// TIA Portal V21 export
// export: Created 2026-10-14T03:09:04.8839945Z, ExportSetting WithDefaults, DisplayName Totally Integrated Automation Portal, DisplayVersion V21, DisplayName STEP 7 Professional, DisplayVersion V21, DisplayName STEP 7 Safety, DisplayVersion V21, DisplayName Tech WebApplication, DisplayVersion V21, DisplayName WinCC Basic/Comfort/Advanced, DisplayVersion V21, DisplayName WinCC Unified, DisplayVersion V21
Screen "10_Startscreen"  800x480, Number=18, Template=01_One_Nav_Level
  on GenerateScreen: GetStartScreenName(); SetTag(Tag := MainNavigationState, Value := 1)
  ScreenLayer 
    Button "Button_12" at 45,392 size 90x32  Mode=Text, TextOff="Place bottle", TextOn="Place bottles"
      VisibilityAnimation "VisibilityAnimation"  RangeEnd=1, RangeStart=1
        tag hmiError
      on Press: ResetBit(Tag := hmiError)
    Rectangle "Rectangle_8" at 682,361 size 88x104  StyleItem=Rectangle
      VisibilityAnimation "VisibilityAnimation"  RangeEnd=1, RangeStart=1
        tag HMI_bottleInfoActive
    GraphicView "Graphic view_4" at 213,87 size 249x237  Picture=Graphic_13
    Button "Button_4" at 45,159 size 90x48  Mode=Text, TextOff="Start", TextOn="Text"
      RangeAppearanceAnimation "RangeAppearanceAnimation"
        tag stateRunning
        0..0: back #404d53, fore #ffffff
      ObjectEnablingAnimation "ObjectEnablingAnimation"
        tag stateRunning
      on Press: SetBit(Tag := hmiStart)
      on Release: ResetBit(Tag := hmiStart)
    Button "Button_5" at 45,215 size 90x48  Mode=Text, TextOff="Stop", TextOn="Text"
      RangeAppearanceAnimation "RangeAppearanceAnimation"
        tag stateRunning
        1..1: back #404d53, fore #ffffff
      ObjectEnablingAnimation "ObjectEnablingAnimation"  RangeEnd=1, RangeStart=1
        tag stateRunning
      on Press: SetBit(Tag := hmiStop)
      on Release: ResetBit(Tag := hmiStop)
    Button "Button_6" at 45,271 size 90x48  Mode=Text, TextOff="Reset", TextOn="Text"
      RangeAppearanceAnimation "RangeAppearanceAnimation"
        tag stateStop
        1..1: back #404d53, fore #ffffff
      ObjectEnablingAnimation "ObjectEnablingAnimation"  RangeEnd=1, RangeStart=1
        tag stateStop
      on Press: SetBit(Tag := hmiReset); ResetBit(Tag := HMI_bottleInfo1); ResetBit(Tag := HMI_bottleInfo2); ResetBit(Tag := HMI_bottleInfo3); ResetBit(Tag := HMI_bottleInfo4); ResetBit(Tag := HMI_bottleInfoActive)
      on Release: ResetBit(Tag := hmiReset)
    IOField "ioKPI" at 700,269 size 68x28  DataFormat=Decimal, FormatPattern=99.9, Mode=Output
      ProcessValue := tankTemperature
    IOField "ioKPI_1" at 687,239 size 76x28  DataFormat=Decimal, FormatPattern=9999, Mode=Output
      ProcessValue := tankLevel
    TextField "Text field_3" at 496,160 size 150x25  Text="Bottles produced"
    Button "Button_1" at 45,354 size 90x32  Mode=Text, TextOff="Next bottle", TextOn="Text"
      ObjectEnablingAnimation "ObjectEnablingAnimation"  RangeEnd=1, RangeStart=1
        tag stateFillingBottle
      RangeAppearanceAnimation "RangeAppearanceAnimation"
        tag stateFillingBottle
        1..1: back #404d53, fore #ffffff
      on Press: SetBit(Tag := hmiNextBottle)
      on Release: ResetBit(Tag := hmiNextBottle)
    TextField "Text field_1" at 610,106 size 150x25  Text="Filling tank"
      VisibilityAnimation "VisibilityAnimation"  Visible=false
        tag stateFillingTank
    TextField "Text field_5" at 496,106 size 49x25  Text="State"
    TextField "Text field_6" at 610,106 size 150x25  Text="Heating tank"
      VisibilityAnimation "VisibilityAnimation"  Visible=false
        tag stateHeatingTank
    TextField "Text field_7" at 610,106 size 150x25  Text="Filling bottle"
      VisibilityAnimation "VisibilityAnimation"  Visible=false
        tag stateFillingBottle
    TextField "Text field_8" at 610,106 size 150x25  Text="Shifting bottle"
      VisibilityAnimation "VisibilityAnimation"  Visible=false
        tag stateShiftingBottle
    TextField "Text field_9" at 610,106 size 150x25  Text="Stop"
      VisibilityAnimation "VisibilityAnimation"  Visible=false
        tag stateStop
    TextField "Text field_10" at 610,106 size 150x25  Text="Reset"
      VisibilityAnimation "VisibilityAnimation"  Visible=false
        tag stateReset
    IOField "ioKPI_2" at 638,160 size 124x28  DataFormat=Decimal, FormatPattern=9999999999, Mode=Output
      ProcessValue := bottlesProduced
    TextField "Text field_11" at 496,191 size 119x25  Text="Bottles faulty"
    IOField "ioKPI_3" at 638,191 size 124x28  DataFormat=Decimal, FormatPattern=9999999999, Mode=Output
      ProcessValue := bootleNumberFaulty
    IOField "ioKPI_4" at 695,329 size 68x28  DataFormat=Decimal, FormatPattern=9.99, Mode=Output
      ProcessValue := bottleLevel
    GraphicView "Graphic view_13" at 326,321 size 17x21  Picture=Graphic_18
    Bar "Bar_1" at 223,115 size 229x206  CountSubDivisions=5, IntegerDigits=3, LargeTickLabelingStep=2, MaximumValue=1600
      RangeAppearanceAnimation "RangeAppearanceAnimation"
        tag tankTemperature
        30..39: back #adaeb5, fore #3f3cff
        40..49: back #adaeb5, fore #4f4dff
        50..59: back #adaeb5, fore #4f4dff
        60..69: back #adaeb5, fore #605eff
        70..72: back #adaeb5, fore #716eff
        73..74: back #adaeb5, fore #8280ff
        75..75: back #adaeb5, fore #9291ff
        76..76: back #adaeb5, fore #9291ff
        77..77: back #adaeb5, fore #a3a2ff
        78..78: back #adaeb5, fore #a3a2ff
        79..79: back #adaeb5, fore #b4b2ff
        80..100: back #adaeb5, fore #b4b2ff
      ProcessValue := tankLevel
    GraphicView "Graphic view_7" at 617,192 size 23x23  Picture=Graphic_58
      VisibilityAnimation "VisibilityAnimation"  RangeEnd=1, RangeStart=1
        tag bottleFaulty
    Rectangle "Rectangle_1" at 238,418 size 32x8  StyleItem=Rectangle
    Rectangle "Rectangle_2" at 199,418 size 32x8  StyleItem=Rectangle
    Line "Line_1" at 200,422 size 266x0  StyleItem=Line
      VisibilityAnimation "VisibilityAnimation"  RangeEnd=2, Visible=false
        tag bottlesProduced
    Rectangle "Rectangle_3" at 279,418 size 32x8  StyleItem=Rectangle
    Rectangle "Rectangle_4" at 317,418 size 32x8  StyleItem=Rectangle
    Rectangle "Rectangle_5" at 356,418 size 32x8  StyleItem=Rectangle
      VisibilityAnimation "VisibilityAnimation"  Visible=false
        tag bottlesProduced
    Rectangle "Rectangle_6" at 396,418 size 32x8  StyleItem=Rectangle
      VisibilityAnimation "VisibilityAnimation"  RangeEnd=1, Visible=false
        tag bottlesProduced
    Rectangle "Rectangle_7" at 436,418 size 32x8  StyleItem=Rectangle
      VisibilityAnimation "VisibilityAnimation"  RangeEnd=2, Visible=false
        tag bottlesProduced
    Line "Line_2" at 200,422 size 225x0  StyleItem=Line
      VisibilityAnimation "VisibilityAnimation"  RangeEnd=1, Visible=false
        tag bottlesProduced
    Line "Line_3" at 200,422 size 185x0  StyleItem=Line
      VisibilityAnimation "VisibilityAnimation"  Visible=false
        tag bottlesProduced
    Line "Line_4" at 201,422 size 147x0  StyleItem=Line
    Button "Button_2" at 322,431 size 26x22  Mode=Graphic, PictureOff=Graphic_50, StyleItem=Button, TextOff="Text", TextOn="Text"
      on Click: SetBit(Tag := HMI_bottleInfo1); ResetBit(Tag := HMI_bottleInfo2); ResetBit(Tag := HMI_bottleInfo3); ResetBit(Tag := HMI_bottleInfo4); HandleBottleInfo()
    Button "Button_7" at 361,431 size 26x22  Mode=Graphic, PictureOff=Graphic_50, StyleItem=Button, TextOff="Text", TextOn="Text"
      VisibilityAnimation "VisibilityAnimation"  Visible=false
        tag bottlesProduced
      on Click: SetBit(Tag := HMI_bottleInfo2); ResetBit(Tag := HMI_bottleInfo1); ResetBit(Tag := HMI_bottleInfo3); ResetBit(Tag := HMI_bottleInfo4); HandleBottleInfo()
    Button "Button_3" at 400,431 size 26x22  Mode=Graphic, PictureOff=Graphic_50, StyleItem=Button, TextOff="Text", TextOn="Text"
      VisibilityAnimation "VisibilityAnimation"  RangeEnd=1, Visible=false
        tag bottlesProduced
      on Click: SetBit(Tag := HMI_bottleInfo3); ResetBit(Tag := HMI_bottleInfo1); ResetBit(Tag := HMI_bottleInfo2); ResetBit(Tag := HMI_bottleInfo4); HandleBottleInfo()
    Button "Button_8" at 440,430 size 26x22  Mode=Graphic, PictureOff=Graphic_50, StyleItem=Button, TextOff="Text", TextOn="Text"
      VisibilityAnimation "VisibilityAnimation"  RangeEnd=2, Visible=false
        tag bottlesProduced
      on Click: SetBit(Tag := HMI_bottleInfo4); ResetBit(Tag := HMI_bottleInfo1); ResetBit(Tag := HMI_bottleInfo2); ResetBit(Tag := HMI_bottleInfo3); HandleBottleInfo()
    IOField "I/O field_1" at 2,459 size 20x20  DataFormat=Binary, FormatPattern=1, Mode=Output
      VisibilityAnimation "VisibilityAnimation"  Visible=false
        tag tempInvisibleObject
      ProcessValue := qrCodeReceived
    GraphicView "Graphic view_1" at 689,384 size 76x76  Picture=QRCode_bottle_one
      VisibilityAnimation "VisibilityAnimation"  RangeEnd=1, RangeStart=1
        tag HMI_bottleInfo1
    TextField "Text field_2" at 666,359 size 78x25  Text="bottle 1"
      VisibilityAnimation "VisibilityAnimation"  RangeEnd=1, RangeStart=1
        tag HMI_bottleInfo1
    TextField "Text field_12" at 665,359 size 78x25  Text="bottle 2"
      VisibilityAnimation "VisibilityAnimation"  RangeEnd=1, RangeStart=1
        tag HMI_bottleInfo2
    GraphicView "Graphic view_3" at 689,384 size 76x76  Picture=QRCode_bottle_two
      VisibilityAnimation "VisibilityAnimation"  RangeEnd=1, RangeStart=1
        tag HMI_bottleInfo2
    TextField "Text field_13" at 666,359 size 78x25  Text="bottle 3"
      VisibilityAnimation "VisibilityAnimation"  RangeEnd=1, RangeStart=1
        tag HMI_bottleInfo3
    TextField "Text field_14" at 665,359 size 78x25  Text="bottle 4"
      VisibilityAnimation "VisibilityAnimation"  RangeEnd=1, RangeStart=1
        tag HMI_bottleInfo4
    GraphicView "Graphic view_5" at 688,384 size 76x76  Picture=QRCode_bottle_three
      VisibilityAnimation "VisibilityAnimation"  RangeEnd=1, RangeStart=1
        tag HMI_bottleInfo3
    GraphicView "Graphic view_6" at 688,386 size 76x76  Picture=QRCode_bottle_four
      VisibilityAnimation "VisibilityAnimation"  RangeEnd=1, RangeStart=1
        tag HMI_bottleInfo4
    Button "Button_10" at 501,392 size 100x32  Mode=Text, PictureOff=Graphic_50, StyleItem=Button, TextOff="Energy data", TextOn="Text"
      on Click: ShowPopupScreen(Name of the screen := EnergyInfo, X coordinate := 0, Y coordinate := 0, Display mode := -1, Animation := -1, Animation speed := 1)
    IOField "ioKPI_6" at 671,299 size 92x28  DataFormat=Decimal, FormatPattern=999.9, Mode=Output
      ProcessValue := tankPressure
    Button "Button_11" at 45,392 size 90x32  Mode=Text, TextOff="Push bottle", TextOn="Place bottles"
      VisibilityAnimation "VisibilityAnimation"
        tag hmiError
      on Press: SetBit(Tag := hmiError)
    GraphicIOField "D6_Pilotlight_Red" at 92,109 size 40x40  Mode=TwoState, OnValue=1, PictureOff=Design_6_PilotLight_Red_Off, PictureOn=Design_6_PilotLight_Red_On
      ProcessValue := stateError
    GraphicIOField "D6_Pilotlight_Green" at 48,109 size 40x40  Mode=TwoState, OnValue=1, PictureOff=Design_6_PilotLight_Green_Off, PictureOn=Design_6_PilotLight_Green_On
      ProcessValue := stateRunning
    TextField "Text field_4" at 610,106 size 150x25  Text="Error"
      VisibilityAnimation "VisibilityAnimation"  Visible=false
        tag stateError
    GraphicView "Graphic view_12" at 138,390 size 28x35  Picture=Graphic_73
    GraphicView "Graphic view_14" at 138,353 size 28x35  Picture=Graphic_74
    TextField "Text field_15" at 496,239 size 113x25  Text="Tank level (l)"
    TextField "Text field_16" at 496,269 size 193x25  Text="Tank temperature (°C)"
    TextField "Text field_17" at 496,299 size 174x25  Text="Tank pressure (hPa)"
    TextField "Text field_18" at 496,329 size 124x25  Text="Bottle level (l)"
    Button "Button_9" at 742,362 size 26x22  Mode=Graphic, PictureOff=Graphic_68, TextOff="Text", TextOn="Text"
      VisibilityAnimation "VisibilityAnimation"  RangeEnd=1, RangeStart=1
        tag HMI_bottleInfoActive
      on Click: ResetBit(Tag := HMI_bottleInfo1); ResetBit(Tag := HMI_bottleInfo2); ResetBit(Tag := HMI_bottleInfo3); ResetBit(Tag := HMI_bottleInfo4); ResetBit(Tag := HMI_bottleInfoActive)
    IOField "I/O field_2" at 23,459 size 20x20  DataFormat=Binary, FormatPattern=1, Mode=Output
      VisibilityAnimation "VisibilityAnimation"  Visible=false
        tag tempInvisibleObject
      ProcessValue := alarmIncoming
    TextField "Text field_19" at 496,132 size 74x25  Text="Batch Id"
    IOField "ioKPI_7" at 638,132 size 124x28  DataFormat=Decimal, FormatPattern=9999999999, Mode=Output
      ProcessValue := batchID
    GraphicView "Graphic view_8" at 318,362 size 36x43  Picture=Graphic_72
      VisibilityAnimation "VisibilityAnimation"  RangeEnd=1, RangeStart=1
        tag hmiError
    GraphicView "bottle finished 1_1" at 279,346 size 30x70  Picture=Graphic_20
    GraphicView "bottle finished 1_2" at 239,346 size 30x70  Picture=Graphic_20
    GraphicView "bottle finished 1_3" at 199,346 size 30x70  Picture=Graphic_20
    GraphicView "bottle finished 1_4" at 357,346 size 30x70  Picture=Graphic_20
      VisibilityAnimation "VisibilityAnimation"  Visible=false
        tag bottlesProduced
    GraphicView "bottle finished 1_5" at 397,346 size 30x70  Picture=Graphic_20
      VisibilityAnimation "VisibilityAnimation"  RangeEnd=1, Visible=false
        tag bottlesProduced
    GraphicView "bottle finished 1_6" at 437,346 size 30x70  Picture=Graphic_20
      VisibilityAnimation "VisibilityAnimation"  RangeEnd=2, Visible=false
        tag bottlesProduced
    Bar "Bar_5" at 443,372 size 20x40  CountSubDivisions=5, IntegerDigits=1, LargeTickLabelingStep=2, MaximumValue=1, MinimumValue=0.01
      VisibilityAnimation "VisibilityAnimation"  RangeEnd=2, Visible=false
        tag bottlesProduced
      ProcessValue := HMI_bottleLevel3
    Bar "Bar_4" at 402,372 size 20x40  CountSubDivisions=5, IntegerDigits=1, LargeTickLabelingStep=2, MaximumValue=1, MinimumValue=0.01
      VisibilityAnimation "VisibilityAnimation"  RangeEnd=1, Visible=false
        tag bottlesProduced
      ProcessValue := HMI_bottleLevel2
    Bar "Bar_3" at 362,372 size 20x40  CountSubDivisions=5, IntegerDigits=1, LargeTickLabelingStep=2, MaximumValue=1, MinimumValue=0.01
      VisibilityAnimation "VisibilityAnimation"  Visible=false
        tag bottlesProduced
      ProcessValue := HMI_bottleLevel1
    GraphicView "bottle finished 1" at 318,346 size 30x70  Picture=Graphic_20
      VisibilityAnimation "VisibilityAnimation"  RangeEnd=1, RangeStart=1, Visible=false
        tag hmiError
    Bar "Bar_2" at 324,371 size 20x40  CountSubDivisions=5, IntegerDigits=1, LargeTickLabelingStep=2, MaximumValue=1, MinimumValue=0.01
      VisibilityAnimation "VisibilityAnimation"  RangeEnd=1, RangeStart=1, Visible=false
        tag hmiError
      ProcessValue := bottleLevel
  ScreenLayer 
    GraphicView "Graphic view_2" at 0,0 size 800x480  Picture=PopUpBackground
      VisibilityAnimation "VisibilityAnimation"  RangeEnd=1, RangeStart=1
        tag PopUpBackground
